Staubli VAL3: MonitorIO1.pgx

program MonitorIO1()
  local bool l_bStopMove
  local bool l_bToHome
  local bool l_bRestartMove
  local bool l_bErr
begin
  l_bRestartMove=true
  l_bStopMove=false
  do
    call io:getDigIO(io:dInput[10],l_bToHome,l_bErr)
    if l_bToHome and (!l_bRestartMove or l_bStopMove)
      l_bRestartMove=true
      l_bStopMove=false
      restartMove()
    endIf

    if !l_bToHome and !l_bStopMove
      l_bStopMove=true
      stopMove()
    endIf

//    if manual:bJogMove
//      if taskStatus("RotGoHome")>=0
//        taskKill("RotGoHome")
//      endIf
//      wait(taskStatus("RotGoHome")<0)

//      stopMove()
//      resetMotion()
//      //2024.11.22 add初始化回零堆栈
//      call ar:resetReturnStack(false)
//      rs:_nOmacStat=9
//      taskKill("Monitor1")
//      wait(taskStatus("Monitor1")<0)
//    endIf
    delay(0)
  until false

end
